Fanuc KAREL source: KA00056.KL

PROGRAM KA00056
%NOLOCKGROUP
VAR
  SRC: POSITION
  DST: JOINTPOS
BEGIN
  DST = SRC
END KA00056
